FUNCTION F_InitializePolarIIChamberServiceStatus : BOOL
VAR_IN_OUT
	ServiceStatus : ST_PolarIIChamber_ServiceStatus;
END_VAR

MEMSET(ADR(ServiceStatus), 0, SIZEOF(ServiceStatus));

// Chamber
F_SetPolarIIChamberServiceIdentity(Status := ServiceStatus.Chamber.SetMode, ServiceId := E_PolarIIChamber_ServiceId.Chamber_SetMode, CompletionBehavior := E_ServiceCompletionBehavior.NaturalCompletion);
F_SetPolarIIChamberServiceIdentity(Status := ServiceStatus.Chamber.Initial, ServiceId := E_PolarIIChamber_ServiceId.Chamber_Initial, CompletionBehavior := E_ServiceCompletionBehavior.NaturalCompletion);
F_SetPolarIIChamberServiceIdentity(Status := ServiceStatus.Chamber.SingleProcess, ServiceId := E_PolarIIChamber_ServiceId.Chamber_SingleProcess, CompletionBehavior := E_ServiceCompletionBehavior.NaturalCompletion);
F_SetPolarIIChamberServiceIdentity(Status := ServiceStatus.Chamber.EMGS, ServiceId := E_PolarIIChamber_ServiceId.Chamber_EMGS, CompletionBehavior := E_ServiceCompletionBehavior.NaturalCompletion);
F_SetPolarIIChamberServiceIdentity(Status := ServiceStatus.Chamber.SetConfig, ServiceId := E_PolarIIChamber_ServiceId.Chamber_SetConfig, CompletionBehavior := E_ServiceCompletionBehavior.NaturalCompletion);
F_SetPolarIIChamberServiceIdentity(Status := ServiceStatus.Chamber.ArmAlignTest, ServiceId := E_PolarIIChamber_ServiceId.Chamber_ArmAlignTest, CompletionBehavior := E_ServiceCompletionBehavior.NaturalCompletion);
F_SetPolarIIChamberServiceIdentity(Status := ServiceStatus.Chamber.ArmTest, ServiceId := E_PolarIIChamber_ServiceId.Chamber_ArmTest, CompletionBehavior := E_ServiceCompletionBehavior.NaturalCompletion);
F_SetPolarIIChamberServiceIdentity(Status := ServiceStatus.Chamber.FlowCalibration, ServiceId := E_PolarIIChamber_ServiceId.Chamber_FlowCalibration, CompletionBehavior := E_ServiceCompletionBehavior.NaturalCompletion);
F_SetPolarIIChamberServiceIdentity(Status := ServiceStatus.Chamber.CupChamberClean, ServiceId := E_PolarIIChamber_ServiceId.Chamber_CupChamberClean, CompletionBehavior := E_ServiceCompletionBehavior.NaturalCompletion);
F_SetPolarIIChamberServiceIdentity(Status := ServiceStatus.Chamber.DoNozzleClean, ServiceId := E_PolarIIChamber_ServiceId.Chamber_DoNozzleClean, CompletionBehavior := E_ServiceCompletionBehavior.NaturalCompletion);
F_SetPolarIIChamberServiceIdentity(Status := ServiceStatus.Chamber.DoNozzlePreflush, ServiceId := E_PolarIIChamber_ServiceId.Chamber_DoNozzlePreflush, CompletionBehavior := E_ServiceCompletionBehavior.NaturalCompletion);

// Arm
F_SetPolarIIChamberServiceIdentity(Status := ServiceStatus.Arm[1].Lift.TopPos, ServiceId := E_PolarIIChamber_ServiceId.Arm1_Lift_TopPos, CompletionBehavior := E_ServiceCompletionBehavior.NaturalCompletion);
F_SetPolarIIChamberServiceIdentity(Status := ServiceStatus.Arm[1].Lift.DownPos, ServiceId := E_PolarIIChamber_ServiceId.Arm1_Lift_DownPos, CompletionBehavior := E_ServiceCompletionBehavior.NaturalCompletion);
F_SetPolarIIChamberServiceIdentity(Status := ServiceStatus.Arm[1].Rotate.JogPositive, ServiceId := E_PolarIIChamber_ServiceId.Arm1_Rotate_JogPositive, CompletionBehavior := E_ServiceCompletionBehavior.ExecuteUntilExternalStop);
F_SetPolarIIChamberServiceIdentity(Status := ServiceStatus.Arm[1].Rotate.JogNegative, ServiceId := E_PolarIIChamber_ServiceId.Arm1_Rotate_JogNegative, CompletionBehavior := E_ServiceCompletionBehavior.ExecuteUntilExternalStop);
F_SetPolarIIChamberServiceIdentity(Status := ServiceStatus.Arm[1].Rotate.IncrementalJog, ServiceId := E_PolarIIChamber_ServiceId.Arm1_Rotate_IncrementalJog, CompletionBehavior := E_ServiceCompletionBehavior.NaturalCompletion);
F_SetPolarIIChamberServiceIdentity(Status := ServiceStatus.Arm[1].Rotate.MoveRecipe, ServiceId := E_PolarIIChamber_ServiceId.Arm1_Rotate_MoveRecipe, CompletionBehavior := E_ServiceCompletionBehavior.NaturalCompletion);
F_SetPolarIIChamberServiceIdentity(Status := ServiceStatus.Arm[1].Rotate.NegLimitPos, ServiceId := E_PolarIIChamber_ServiceId.Arm1_Rotate_NegLimitPos, CompletionBehavior := E_ServiceCompletionBehavior.NaturalCompletion);
F_SetPolarIIChamberServiceIdentity(Status := ServiceStatus.Arm[1].Rotate.PosLimitPos, ServiceId := E_PolarIIChamber_ServiceId.Arm1_Rotate_PosLimitPos, CompletionBehavior := E_ServiceCompletionBehavior.NaturalCompletion);
F_SetPolarIIChamberServiceIdentity(Status := ServiceStatus.Arm[1].Rotate.NozzlePortPos, ServiceId := E_PolarIIChamber_ServiceId.Arm1_Rotate_NozPortPos, CompletionBehavior := E_ServiceCompletionBehavior.NaturalCompletion);
F_SetPolarIIChamberServiceIdentity(Status := ServiceStatus.Arm[1].Rotate.Noz1CenterPos, ServiceId := E_PolarIIChamber_ServiceId.Arm1_Rotate_Noz1CenterPos, CompletionBehavior := E_ServiceCompletionBehavior.NaturalCompletion);
F_SetPolarIIChamberServiceIdentity(Status := ServiceStatus.Arm[1].Rotate.Noz2CenterPos, ServiceId := E_PolarIIChamber_ServiceId.Arm1_Rotate_Noz2CenterPos, CompletionBehavior := E_ServiceCompletionBehavior.NaturalCompletion);
F_SetPolarIIChamberServiceIdentity(Status := ServiceStatus.Arm[1].Rotate.Noz3CenterPos, ServiceId := E_PolarIIChamber_ServiceId.Arm1_Rotate_Noz3CenterPos, CompletionBehavior := E_ServiceCompletionBehavior.NaturalCompletion);
F_SetPolarIIChamberServiceIdentity(Status := ServiceStatus.Arm[1].Nozzle[1].ChemicalSupply, ServiceId := E_PolarIIChamber_ServiceId.Arm1_Noz1_ChemicalSupply, CompletionBehavior := E_ServiceCompletionBehavior.ExecuteUntilExternalStop);
F_SetPolarIIChamberServiceIdentity(Status := ServiceStatus.Arm[1].Nozzle[2].ChemicalSupply, ServiceId := E_PolarIIChamber_ServiceId.Arm1_Noz2_ChemicalSupply, CompletionBehavior := E_ServiceCompletionBehavior.ExecuteUntilExternalStop);
F_SetPolarIIChamberServiceIdentity(Status := ServiceStatus.Arm[1].Nozzle[3].ChemicalSupply, ServiceId := E_PolarIIChamber_ServiceId.Arm1_Noz3_ChemicalSupply, CompletionBehavior := E_ServiceCompletionBehavior.ExecuteUntilExternalStop);
F_SetPolarIIChamberServiceIdentity(Status := ServiceStatus.Arm[1].NozzlePort.Nozzle[1].Supply, ServiceId := E_PolarIIChamber_ServiceId.Arm1_NozPortNoz1_Supply, CompletionBehavior := E_ServiceCompletionBehavior.ExecuteUntilExternalStop);
F_SetPolarIIChamberServiceIdentity(Status := ServiceStatus.Arm[1].NozzlePort.Nozzle[2].Supply, ServiceId := E_PolarIIChamber_ServiceId.Arm1_NozPortNoz2_Supply, CompletionBehavior := E_ServiceCompletionBehavior.ExecuteUntilExternalStop);
F_SetPolarIIChamberServiceIdentity(Status := ServiceStatus.Arm[1].NozzlePort.Nozzle[3].Supply, ServiceId := E_PolarIIChamber_ServiceId.Arm1_NozPortNoz3_Supply, CompletionBehavior := E_ServiceCompletionBehavior.ExecuteUntilExternalStop);
F_SetPolarIIChamberServiceIdentity(Status := ServiceStatus.Arm[1].NozzlePort.DrainSelect1, ServiceId := E_PolarIIChamber_ServiceId.Arm1_NozPortDrainer_Select1, CompletionBehavior := E_ServiceCompletionBehavior.NaturalCompletion);
F_SetPolarIIChamberServiceIdentity(Status := ServiceStatus.Arm[1].NozzlePort.DrainSelect2, ServiceId := E_PolarIIChamber_ServiceId.Arm1_NozPortDrainer_Select2, CompletionBehavior := E_ServiceCompletionBehavior.NaturalCompletion);
F_SetPolarIIChamberServiceIdentity(Status := ServiceStatus.Arm[1].NozzlePort.DrainSelect3, ServiceId := E_PolarIIChamber_ServiceId.Arm1_NozPortDrainer_Select3, CompletionBehavior := E_ServiceCompletionBehavior.NaturalCompletion);
F_SetPolarIIChamberServiceIdentity(Status := ServiceStatus.Arm[2].Lift.TopPos, ServiceId := E_PolarIIChamber_ServiceId.Arm2_Lift_TopPos, CompletionBehavior := E_ServiceCompletionBehavior.NaturalCompletion);
F_SetPolarIIChamberServiceIdentity(Status := ServiceStatus.Arm[2].Lift.DownPos, ServiceId := E_PolarIIChamber_ServiceId.Arm2_Lift_DownPos, CompletionBehavior := E_ServiceCompletionBehavior.NaturalCompletion);
F_SetPolarIIChamberServiceIdentity(Status := ServiceStatus.Arm[2].Rotate.JogPositive, ServiceId := E_PolarIIChamber_ServiceId.Arm2_Rotate_JogPositive, CompletionBehavior := E_ServiceCompletionBehavior.ExecuteUntilExternalStop);
F_SetPolarIIChamberServiceIdentity(Status := ServiceStatus.Arm[2].Rotate.JogNegative, ServiceId := E_PolarIIChamber_ServiceId.Arm2_Rotate_JogNegative, CompletionBehavior := E_ServiceCompletionBehavior.ExecuteUntilExternalStop);
F_SetPolarIIChamberServiceIdentity(Status := ServiceStatus.Arm[2].Rotate.IncrementalJog, ServiceId := E_PolarIIChamber_ServiceId.Arm2_Rotate_IncrementalJog, CompletionBehavior := E_ServiceCompletionBehavior.NaturalCompletion);
F_SetPolarIIChamberServiceIdentity(Status := ServiceStatus.Arm[2].Rotate.MoveRecipe, ServiceId := E_PolarIIChamber_ServiceId.Arm2_Rotate_MoveRecipe, CompletionBehavior := E_ServiceCompletionBehavior.NaturalCompletion);
F_SetPolarIIChamberServiceIdentity(Status := ServiceStatus.Arm[2].Rotate.NegLimitPos, ServiceId := E_PolarIIChamber_ServiceId.Arm2_Rotate_NegLimitPos, CompletionBehavior := E_ServiceCompletionBehavior.NaturalCompletion);
F_SetPolarIIChamberServiceIdentity(Status := ServiceStatus.Arm[2].Rotate.PosLimitPos, ServiceId := E_PolarIIChamber_ServiceId.Arm2_Rotate_PosLimitPos, CompletionBehavior := E_ServiceCompletionBehavior.NaturalCompletion);
F_SetPolarIIChamberServiceIdentity(Status := ServiceStatus.Arm[2].Rotate.NozzlePortPos, ServiceId := E_PolarIIChamber_ServiceId.Arm2_Rotate_NozPortPos, CompletionBehavior := E_ServiceCompletionBehavior.NaturalCompletion);
F_SetPolarIIChamberServiceIdentity(Status := ServiceStatus.Arm[2].Rotate.Noz1CenterPos, ServiceId := E_PolarIIChamber_ServiceId.Arm2_Rotate_Noz1CenterPos, CompletionBehavior := E_ServiceCompletionBehavior.NaturalCompletion);
F_SetPolarIIChamberServiceIdentity(Status := ServiceStatus.Arm[2].Rotate.Noz2CenterPos, ServiceId := E_PolarIIChamber_ServiceId.Arm2_Rotate_Noz2CenterPos, CompletionBehavior := E_ServiceCompletionBehavior.NaturalCompletion);
F_SetPolarIIChamberServiceIdentity(Status := ServiceStatus.Arm[2].Rotate.Noz3CenterPos, ServiceId := E_PolarIIChamber_ServiceId.Arm2_Rotate_Noz3CenterPos, CompletionBehavior := E_ServiceCompletionBehavior.NaturalCompletion);
F_SetPolarIIChamberServiceIdentity(Status := ServiceStatus.Arm[2].Nozzle[1].ChemicalSupply, ServiceId := E_PolarIIChamber_ServiceId.Arm2_Noz1_ChemicalSupply, CompletionBehavior := E_ServiceCompletionBehavior.ExecuteUntilExternalStop);
F_SetPolarIIChamberServiceIdentity(Status := ServiceStatus.Arm[2].Nozzle[2].ChemicalSupply, ServiceId := E_PolarIIChamber_ServiceId.Arm2_Noz2_ChemicalSupply, CompletionBehavior := E_ServiceCompletionBehavior.ExecuteUntilExternalStop);
F_SetPolarIIChamberServiceIdentity(Status := ServiceStatus.Arm[2].Nozzle[3].ChemicalSupply, ServiceId := E_PolarIIChamber_ServiceId.Arm2_Noz3_ChemicalSupply, CompletionBehavior := E_ServiceCompletionBehavior.ExecuteUntilExternalStop);
F_SetPolarIIChamberServiceIdentity(Status := ServiceStatus.Arm[2].NozzlePort.Nozzle[1].Supply, ServiceId := E_PolarIIChamber_ServiceId.Arm2_NozPortNoz1_Supply, CompletionBehavior := E_ServiceCompletionBehavior.ExecuteUntilExternalStop);
F_SetPolarIIChamberServiceIdentity(Status := ServiceStatus.Arm[2].NozzlePort.Nozzle[2].Supply, ServiceId := E_PolarIIChamber_ServiceId.Arm2_NozPortNoz2_Supply, CompletionBehavior := E_ServiceCompletionBehavior.ExecuteUntilExternalStop);
F_SetPolarIIChamberServiceIdentity(Status := ServiceStatus.Arm[2].NozzlePort.Nozzle[3].Supply, ServiceId := E_PolarIIChamber_ServiceId.Arm2_NozPortNoz3_Supply, CompletionBehavior := E_ServiceCompletionBehavior.ExecuteUntilExternalStop);
F_SetPolarIIChamberServiceIdentity(Status := ServiceStatus.Arm[2].NozzlePort.DrainSelect1, ServiceId := E_PolarIIChamber_ServiceId.Arm2_NozPortDrainer_Select1, CompletionBehavior := E_ServiceCompletionBehavior.NaturalCompletion);
F_SetPolarIIChamberServiceIdentity(Status := ServiceStatus.Arm[2].NozzlePort.DrainSelect2, ServiceId := E_PolarIIChamber_ServiceId.Arm2_NozPortDrainer_Select2, CompletionBehavior := E_ServiceCompletionBehavior.NaturalCompletion);
F_SetPolarIIChamberServiceIdentity(Status := ServiceStatus.Arm[2].NozzlePort.DrainSelect3, ServiceId := E_PolarIIChamber_ServiceId.Arm2_NozPortDrainer_Select3, CompletionBehavior := E_ServiceCompletionBehavior.NaturalCompletion);
F_SetPolarIIChamberServiceIdentity(Status := ServiceStatus.Arm[3].Lift.TopPos, ServiceId := E_PolarIIChamber_ServiceId.Arm3_Lift_TopPos, CompletionBehavior := E_ServiceCompletionBehavior.NaturalCompletion);
F_SetPolarIIChamberServiceIdentity(Status := ServiceStatus.Arm[3].Lift.DownPos, ServiceId := E_PolarIIChamber_ServiceId.Arm3_Lift_DownPos, CompletionBehavior := E_ServiceCompletionBehavior.NaturalCompletion);
F_SetPolarIIChamberServiceIdentity(Status := ServiceStatus.Arm[3].Rotate.JogPositive, ServiceId := E_PolarIIChamber_ServiceId.Arm3_Rotate_JogPositive, CompletionBehavior := E_ServiceCompletionBehavior.ExecuteUntilExternalStop);
F_SetPolarIIChamberServiceIdentity(Status := ServiceStatus.Arm[3].Rotate.JogNegative, ServiceId := E_PolarIIChamber_ServiceId.Arm3_Rotate_JogNegative, CompletionBehavior := E_ServiceCompletionBehavior.ExecuteUntilExternalStop);
F_SetPolarIIChamberServiceIdentity(Status := ServiceStatus.Arm[3].Rotate.IncrementalJog, ServiceId := E_PolarIIChamber_ServiceId.Arm3_Rotate_IncrementalJog, CompletionBehavior := E_ServiceCompletionBehavior.NaturalCompletion);
F_SetPolarIIChamberServiceIdentity(Status := ServiceStatus.Arm[3].Rotate.MoveRecipe, ServiceId := E_PolarIIChamber_ServiceId.Arm3_Rotate_MoveRecipe, CompletionBehavior := E_ServiceCompletionBehavior.NaturalCompletion);
F_SetPolarIIChamberServiceIdentity(Status := ServiceStatus.Arm[3].Rotate.NegLimitPos, ServiceId := E_PolarIIChamber_ServiceId.Arm3_Rotate_NegLimitPos, CompletionBehavior := E_ServiceCompletionBehavior.NaturalCompletion);
F_SetPolarIIChamberServiceIdentity(Status := ServiceStatus.Arm[3].Rotate.PosLimitPos, ServiceId := E_PolarIIChamber_ServiceId.Arm3_Rotate_PosLimitPos, CompletionBehavior := E_ServiceCompletionBehavior.NaturalCompletion);
F_SetPolarIIChamberServiceIdentity(Status := ServiceStatus.Arm[3].Rotate.Noz1CenterPos, ServiceId := E_PolarIIChamber_ServiceId.Arm3_Rotate_Noz1CenterPos, CompletionBehavior := E_ServiceCompletionBehavior.NaturalCompletion);
F_SetPolarIIChamberServiceIdentity(Status := ServiceStatus.Arm[3].Rotate.Noz2CenterPos, ServiceId := E_PolarIIChamber_ServiceId.Arm3_Rotate_Noz2CenterPos, CompletionBehavior := E_ServiceCompletionBehavior.NaturalCompletion);
F_SetPolarIIChamberServiceIdentity(Status := ServiceStatus.Arm[3].Nozzle[1].ChemicalSupply, ServiceId := E_PolarIIChamber_ServiceId.Arm3_Noz1_ChemicalSupply, CompletionBehavior := E_ServiceCompletionBehavior.ExecuteUntilExternalStop);
F_SetPolarIIChamberServiceIdentity(Status := ServiceStatus.Arm[3].Nozzle[2].ChemicalSupply, ServiceId := E_PolarIIChamber_ServiceId.Arm3_Noz2_ChemicalSupply, CompletionBehavior := E_ServiceCompletionBehavior.ExecuteUntilExternalStop);
// Arm[3] has no third nozzle or nozzle port. Keep ServiceId = 0, but provide
// CompletionBehavior so the current SDK STRUCT scanner can complete validation.
ServiceStatus.Arm[3].Rotate.NozzlePortPos.CompletionBehavior := E_ServiceCompletionBehavior.NaturalCompletion;
ServiceStatus.Arm[3].Rotate.Noz3CenterPos.CompletionBehavior := E_ServiceCompletionBehavior.NaturalCompletion;
ServiceStatus.Arm[3].Nozzle[3].ChemicalSupply.CompletionBehavior := E_ServiceCompletionBehavior.ExecuteUntilExternalStop;
ServiceStatus.Arm[3].NozzlePort.Nozzle[1].Supply.CompletionBehavior := E_ServiceCompletionBehavior.ExecuteUntilExternalStop;
ServiceStatus.Arm[3].NozzlePort.Nozzle[2].Supply.CompletionBehavior := E_ServiceCompletionBehavior.ExecuteUntilExternalStop;
ServiceStatus.Arm[3].NozzlePort.Nozzle[3].Supply.CompletionBehavior := E_ServiceCompletionBehavior.ExecuteUntilExternalStop;
ServiceStatus.Arm[3].NozzlePort.DrainSelect1.CompletionBehavior := E_ServiceCompletionBehavior.NaturalCompletion;
ServiceStatus.Arm[3].NozzlePort.DrainSelect2.CompletionBehavior := E_ServiceCompletionBehavior.NaturalCompletion;
ServiceStatus.Arm[3].NozzlePort.DrainSelect3.CompletionBehavior := E_ServiceCompletionBehavior.NaturalCompletion;
F_SetPolarIIChamberServiceIdentity(Status := ServiceStatus.Arm[4].Lift.TopPos, ServiceId := E_PolarIIChamber_ServiceId.Arm4_Lift_TopPos, CompletionBehavior := E_ServiceCompletionBehavior.NaturalCompletion);
F_SetPolarIIChamberServiceIdentity(Status := ServiceStatus.Arm[4].Lift.DownPos, ServiceId := E_PolarIIChamber_ServiceId.Arm4_Lift_DownPos, CompletionBehavior := E_ServiceCompletionBehavior.NaturalCompletion);
F_SetPolarIIChamberServiceIdentity(Status := ServiceStatus.Arm[4].Rotate.JogPositive, ServiceId := E_PolarIIChamber_ServiceId.Arm4_Rotate_JogPositive, CompletionBehavior := E_ServiceCompletionBehavior.ExecuteUntilExternalStop);
F_SetPolarIIChamberServiceIdentity(Status := ServiceStatus.Arm[4].Rotate.JogNegative, ServiceId := E_PolarIIChamber_ServiceId.Arm4_Rotate_JogNegative, CompletionBehavior := E_ServiceCompletionBehavior.ExecuteUntilExternalStop);
F_SetPolarIIChamberServiceIdentity(Status := ServiceStatus.Arm[4].Rotate.IncrementalJog, ServiceId := E_PolarIIChamber_ServiceId.Arm4_Rotate_IncrementalJog, CompletionBehavior := E_ServiceCompletionBehavior.NaturalCompletion);
F_SetPolarIIChamberServiceIdentity(Status := ServiceStatus.Arm[4].Rotate.MoveRecipe, ServiceId := E_PolarIIChamber_ServiceId.Arm4_Rotate_MoveRecipe, CompletionBehavior := E_ServiceCompletionBehavior.NaturalCompletion);
F_SetPolarIIChamberServiceIdentity(Status := ServiceStatus.Arm[4].Rotate.NegLimitPos, ServiceId := E_PolarIIChamber_ServiceId.Arm4_Rotate_NegLimitPos, CompletionBehavior := E_ServiceCompletionBehavior.NaturalCompletion);
F_SetPolarIIChamberServiceIdentity(Status := ServiceStatus.Arm[4].Rotate.PosLimitPos, ServiceId := E_PolarIIChamber_ServiceId.Arm4_Rotate_PosLimitPos, CompletionBehavior := E_ServiceCompletionBehavior.NaturalCompletion);
F_SetPolarIIChamberServiceIdentity(Status := ServiceStatus.Arm[4].Rotate.Noz1CenterPos, ServiceId := E_PolarIIChamber_ServiceId.Arm4_Rotate_Noz1CenterPos, CompletionBehavior := E_ServiceCompletionBehavior.NaturalCompletion);
F_SetPolarIIChamberServiceIdentity(Status := ServiceStatus.Arm[4].Nozzle[1].ChemicalSupply, ServiceId := E_PolarIIChamber_ServiceId.Arm4_Noz1_ChemicalSupply, CompletionBehavior := E_ServiceCompletionBehavior.ExecuteUntilExternalStop);
// Arm[4] has no second/third nozzle or nozzle port. Keep ServiceId = 0, but
// provide CompletionBehavior for compatibility with the current SDK scanner.
ServiceStatus.Arm[4].Rotate.NozzlePortPos.CompletionBehavior := E_ServiceCompletionBehavior.NaturalCompletion;
ServiceStatus.Arm[4].Rotate.Noz2CenterPos.CompletionBehavior := E_ServiceCompletionBehavior.NaturalCompletion;
ServiceStatus.Arm[4].Rotate.Noz3CenterPos.CompletionBehavior := E_ServiceCompletionBehavior.NaturalCompletion;
ServiceStatus.Arm[4].Nozzle[2].ChemicalSupply.CompletionBehavior := E_ServiceCompletionBehavior.ExecuteUntilExternalStop;
ServiceStatus.Arm[4].Nozzle[3].ChemicalSupply.CompletionBehavior := E_ServiceCompletionBehavior.ExecuteUntilExternalStop;
ServiceStatus.Arm[4].NozzlePort.Nozzle[1].Supply.CompletionBehavior := E_ServiceCompletionBehavior.ExecuteUntilExternalStop;
ServiceStatus.Arm[4].NozzlePort.Nozzle[2].Supply.CompletionBehavior := E_ServiceCompletionBehavior.ExecuteUntilExternalStop;
ServiceStatus.Arm[4].NozzlePort.Nozzle[3].Supply.CompletionBehavior := E_ServiceCompletionBehavior.ExecuteUntilExternalStop;
ServiceStatus.Arm[4].NozzlePort.DrainSelect1.CompletionBehavior := E_ServiceCompletionBehavior.NaturalCompletion;
ServiceStatus.Arm[4].NozzlePort.DrainSelect2.CompletionBehavior := E_ServiceCompletionBehavior.NaturalCompletion;
ServiceStatus.Arm[4].NozzlePort.DrainSelect3.CompletionBehavior := E_ServiceCompletionBehavior.NaturalCompletion;

// Cup
F_SetPolarIIChamberServiceIdentity(Status := ServiceStatus.Cup[1].Lift.JogPositive, ServiceId := E_PolarIIChamber_ServiceId.Cup1_Lift_JogPositive, CompletionBehavior := E_ServiceCompletionBehavior.ExecuteUntilExternalStop);
F_SetPolarIIChamberServiceIdentity(Status := ServiceStatus.Cup[1].Lift.JogNegative, ServiceId := E_PolarIIChamber_ServiceId.Cup1_Lift_JogNegative, CompletionBehavior := E_ServiceCompletionBehavior.ExecuteUntilExternalStop);
F_SetPolarIIChamberServiceIdentity(Status := ServiceStatus.Cup[1].Lift.IncrementalJog, ServiceId := E_PolarIIChamber_ServiceId.Cup1_Lift_IncrementalJog, CompletionBehavior := E_ServiceCompletionBehavior.NaturalCompletion);
F_SetPolarIIChamberServiceIdentity(Status := ServiceStatus.Cup[1].Lift.DecoupleStop, ServiceId := E_PolarIIChamber_ServiceId.Cup1_Lift_DecoupleStop, CompletionBehavior := E_ServiceCompletionBehavior.NaturalCompletion);
F_SetPolarIIChamberServiceIdentity(Status := ServiceStatus.Cup[1].Lift.TopPos, ServiceId := E_PolarIIChamber_ServiceId.Cup1_Lift_TopPos, CompletionBehavior := E_ServiceCompletionBehavior.NaturalCompletion);
F_SetPolarIIChamberServiceIdentity(Status := ServiceStatus.Cup[1].Lift.MiddlePos, ServiceId := E_PolarIIChamber_ServiceId.Cup1_Lift_MiddlePos, CompletionBehavior := E_ServiceCompletionBehavior.NaturalCompletion);
F_SetPolarIIChamberServiceIdentity(Status := ServiceStatus.Cup[1].Lift.DownPos, ServiceId := E_PolarIIChamber_ServiceId.Cup1_Lift_DownPos, CompletionBehavior := E_ServiceCompletionBehavior.NaturalCompletion);
F_SetPolarIIChamberServiceIdentity(Status := ServiceStatus.Cup[1].Drainer.Select1, ServiceId := E_PolarIIChamber_ServiceId.Cup1_Drainer_Select1, CompletionBehavior := E_ServiceCompletionBehavior.NaturalCompletion);
F_SetPolarIIChamberServiceIdentity(Status := ServiceStatus.Cup[1].Drainer.Select2, ServiceId := E_PolarIIChamber_ServiceId.Cup1_Drainer_Select2, CompletionBehavior := E_ServiceCompletionBehavior.NaturalCompletion);
F_SetPolarIIChamberServiceIdentity(Status := ServiceStatus.Cup[1].Drainer.Select3, ServiceId := E_PolarIIChamber_ServiceId.Cup1_Drainer_Select3, CompletionBehavior := E_ServiceCompletionBehavior.NaturalCompletion);
F_SetPolarIIChamberServiceIdentity(Status := ServiceStatus.Cup[2].Lift.JogPositive, ServiceId := E_PolarIIChamber_ServiceId.Cup2_Lift_JogPositive, CompletionBehavior := E_ServiceCompletionBehavior.ExecuteUntilExternalStop);
F_SetPolarIIChamberServiceIdentity(Status := ServiceStatus.Cup[2].Lift.JogNegative, ServiceId := E_PolarIIChamber_ServiceId.Cup2_Lift_JogNegative, CompletionBehavior := E_ServiceCompletionBehavior.ExecuteUntilExternalStop);
F_SetPolarIIChamberServiceIdentity(Status := ServiceStatus.Cup[2].Lift.IncrementalJog, ServiceId := E_PolarIIChamber_ServiceId.Cup2_Lift_IncrementalJog, CompletionBehavior := E_ServiceCompletionBehavior.NaturalCompletion);
F_SetPolarIIChamberServiceIdentity(Status := ServiceStatus.Cup[2].Lift.DecoupleStop, ServiceId := E_PolarIIChamber_ServiceId.Cup2_Lift_DecoupleStop, CompletionBehavior := E_ServiceCompletionBehavior.NaturalCompletion);
F_SetPolarIIChamberServiceIdentity(Status := ServiceStatus.Cup[2].Lift.TopPos, ServiceId := E_PolarIIChamber_ServiceId.Cup2_Lift_TopPos, CompletionBehavior := E_ServiceCompletionBehavior.NaturalCompletion);
F_SetPolarIIChamberServiceIdentity(Status := ServiceStatus.Cup[2].Lift.MiddlePos, ServiceId := E_PolarIIChamber_ServiceId.Cup2_Lift_MiddlePos, CompletionBehavior := E_ServiceCompletionBehavior.NaturalCompletion);
F_SetPolarIIChamberServiceIdentity(Status := ServiceStatus.Cup[2].Lift.DownPos, ServiceId := E_PolarIIChamber_ServiceId.Cup2_Lift_DownPos, CompletionBehavior := E_ServiceCompletionBehavior.NaturalCompletion);
F_SetPolarIIChamberServiceIdentity(Status := ServiceStatus.Cup[2].Drainer.Select1, ServiceId := E_PolarIIChamber_ServiceId.Cup2_Drainer_Select1, CompletionBehavior := E_ServiceCompletionBehavior.NaturalCompletion);
F_SetPolarIIChamberServiceIdentity(Status := ServiceStatus.Cup[2].Drainer.Select2, ServiceId := E_PolarIIChamber_ServiceId.Cup2_Drainer_Select2, CompletionBehavior := E_ServiceCompletionBehavior.NaturalCompletion);
F_SetPolarIIChamberServiceIdentity(Status := ServiceStatus.Cup[2].Drainer.Select3, ServiceId := E_PolarIIChamber_ServiceId.Cup2_Drainer_Select3, CompletionBehavior := E_ServiceCompletionBehavior.NaturalCompletion);
F_SetPolarIIChamberServiceIdentity(Status := ServiceStatus.Cup[3].Lift.JogPositive, ServiceId := E_PolarIIChamber_ServiceId.Cup3_Lift_JogPositive, CompletionBehavior := E_ServiceCompletionBehavior.ExecuteUntilExternalStop);
F_SetPolarIIChamberServiceIdentity(Status := ServiceStatus.Cup[3].Lift.JogNegative, ServiceId := E_PolarIIChamber_ServiceId.Cup3_Lift_JogNegative, CompletionBehavior := E_ServiceCompletionBehavior.ExecuteUntilExternalStop);
F_SetPolarIIChamberServiceIdentity(Status := ServiceStatus.Cup[3].Lift.IncrementalJog, ServiceId := E_PolarIIChamber_ServiceId.Cup3_Lift_IncrementalJog, CompletionBehavior := E_ServiceCompletionBehavior.NaturalCompletion);
F_SetPolarIIChamberServiceIdentity(Status := ServiceStatus.Cup[3].Lift.DecoupleStop, ServiceId := E_PolarIIChamber_ServiceId.Cup3_Lift_DecoupleStop, CompletionBehavior := E_ServiceCompletionBehavior.NaturalCompletion);
F_SetPolarIIChamberServiceIdentity(Status := ServiceStatus.Cup[3].Lift.TopPos, ServiceId := E_PolarIIChamber_ServiceId.Cup3_Lift_TopPos, CompletionBehavior := E_ServiceCompletionBehavior.NaturalCompletion);
F_SetPolarIIChamberServiceIdentity(Status := ServiceStatus.Cup[3].Lift.MiddlePos, ServiceId := E_PolarIIChamber_ServiceId.Cup3_Lift_MiddlePos, CompletionBehavior := E_ServiceCompletionBehavior.NaturalCompletion);
F_SetPolarIIChamberServiceIdentity(Status := ServiceStatus.Cup[3].Lift.DownPos, ServiceId := E_PolarIIChamber_ServiceId.Cup3_Lift_DownPos, CompletionBehavior := E_ServiceCompletionBehavior.NaturalCompletion);
F_SetPolarIIChamberServiceIdentity(Status := ServiceStatus.Cup[3].Drainer.Select1, ServiceId := E_PolarIIChamber_ServiceId.Cup3_Drainer_Select1, CompletionBehavior := E_ServiceCompletionBehavior.NaturalCompletion);
F_SetPolarIIChamberServiceIdentity(Status := ServiceStatus.Cup[3].Drainer.Select2, ServiceId := E_PolarIIChamber_ServiceId.Cup3_Drainer_Select2, CompletionBehavior := E_ServiceCompletionBehavior.NaturalCompletion);
F_SetPolarIIChamberServiceIdentity(Status := ServiceStatus.Cup[3].Drainer.Select3, ServiceId := E_PolarIIChamber_ServiceId.Cup3_Drainer_Select3, CompletionBehavior := E_ServiceCompletionBehavior.NaturalCompletion);
F_SetPolarIIChamberServiceIdentity(Status := ServiceStatus.Cup[4].Lift.JogPositive, ServiceId := E_PolarIIChamber_ServiceId.Cup4_Lift_JogPositive, CompletionBehavior := E_ServiceCompletionBehavior.ExecuteUntilExternalStop);
F_SetPolarIIChamberServiceIdentity(Status := ServiceStatus.Cup[4].Lift.JogNegative, ServiceId := E_PolarIIChamber_ServiceId.Cup4_Lift_JogNegative, CompletionBehavior := E_ServiceCompletionBehavior.ExecuteUntilExternalStop);
F_SetPolarIIChamberServiceIdentity(Status := ServiceStatus.Cup[4].Lift.IncrementalJog, ServiceId := E_PolarIIChamber_ServiceId.Cup4_Lift_IncrementalJog, CompletionBehavior := E_ServiceCompletionBehavior.NaturalCompletion);
F_SetPolarIIChamberServiceIdentity(Status := ServiceStatus.Cup[4].Lift.DecoupleStop, ServiceId := E_PolarIIChamber_ServiceId.Cup4_Lift_DecoupleStop, CompletionBehavior := E_ServiceCompletionBehavior.NaturalCompletion);
F_SetPolarIIChamberServiceIdentity(Status := ServiceStatus.Cup[4].Lift.TopPos, ServiceId := E_PolarIIChamber_ServiceId.Cup4_Lift_TopPos, CompletionBehavior := E_ServiceCompletionBehavior.NaturalCompletion);
F_SetPolarIIChamberServiceIdentity(Status := ServiceStatus.Cup[4].Lift.MiddlePos, ServiceId := E_PolarIIChamber_ServiceId.Cup4_Lift_MiddlePos, CompletionBehavior := E_ServiceCompletionBehavior.NaturalCompletion);
F_SetPolarIIChamberServiceIdentity(Status := ServiceStatus.Cup[4].Lift.DownPos, ServiceId := E_PolarIIChamber_ServiceId.Cup4_Lift_DownPos, CompletionBehavior := E_ServiceCompletionBehavior.NaturalCompletion);
F_SetPolarIIChamberServiceIdentity(Status := ServiceStatus.Cup[4].Drainer.Select1, ServiceId := E_PolarIIChamber_ServiceId.Cup4_Drainer_Select1, CompletionBehavior := E_ServiceCompletionBehavior.NaturalCompletion);
F_SetPolarIIChamberServiceIdentity(Status := ServiceStatus.Cup[4].Drainer.Select2, ServiceId := E_PolarIIChamber_ServiceId.Cup4_Drainer_Select2, CompletionBehavior := E_ServiceCompletionBehavior.NaturalCompletion);
F_SetPolarIIChamberServiceIdentity(Status := ServiceStatus.Cup[4].Drainer.Select3, ServiceId := E_PolarIIChamber_ServiceId.Cup4_Drainer_Select3, CompletionBehavior := E_ServiceCompletionBehavior.NaturalCompletion);

// Holder
F_SetPolarIIChamberServiceIdentity(Status := ServiceStatus.Holder.Gripper.Open, ServiceId := E_PolarIIChamber_ServiceId.Holder_Gripper_Open, CompletionBehavior := E_ServiceCompletionBehavior.NaturalCompletion);
F_SetPolarIIChamberServiceIdentity(Status := ServiceStatus.Holder.Gripper.Close, ServiceId := E_PolarIIChamber_ServiceId.Holder_Gripper_Close, CompletionBehavior := E_ServiceCompletionBehavior.NaturalCompletion);
F_SetPolarIIChamberServiceIdentity(Status := ServiceStatus.Holder.Rotate.OPR, ServiceId := E_PolarIIChamber_ServiceId.Holder_Rotate_OPR, CompletionBehavior := E_ServiceCompletionBehavior.NaturalCompletion);
F_SetPolarIIChamberServiceIdentity(Status := ServiceStatus.Holder.Rotate.MoveVelocityCW, ServiceId := E_PolarIIChamber_ServiceId.Holder_Rotate_MoveVelocityCW, CompletionBehavior := E_ServiceCompletionBehavior.ExecuteUntilExternalStop);
F_SetPolarIIChamberServiceIdentity(Status := ServiceStatus.Holder.Rotate.MoveVelocityCCW, ServiceId := E_PolarIIChamber_ServiceId.Holder_Rotate_MoveVelocityCCW, CompletionBehavior := E_ServiceCompletionBehavior.ExecuteUntilExternalStop);
F_SetPolarIIChamberServiceIdentity(Status := ServiceStatus.Holder.Rotate.MoveModulo, ServiceId := E_PolarIIChamber_ServiceId.Holder_Rotate_MoveModulo, CompletionBehavior := E_ServiceCompletionBehavior.NaturalCompletion);
F_SetPolarIIChamberServiceIdentity(Status := ServiceStatus.Holder.VacuumEstablish, ServiceId := E_PolarIIChamber_ServiceId.Holder_VacuumEstablish, CompletionBehavior := E_ServiceCompletionBehavior.ExecuteUntilExternalStop);

// FixedNozzle
F_SetPolarIIChamberServiceIdentity(Status := ServiceStatus.FixedNozzle[1].ChemicalSupply, ServiceId := E_PolarIIChamber_ServiceId.FixedNoz1_ChemicalSupply, CompletionBehavior := E_ServiceCompletionBehavior.ExecuteUntilExternalStop);
F_SetPolarIIChamberServiceIdentity(Status := ServiceStatus.FixedNozzle[2].ChemicalSupply, ServiceId := E_PolarIIChamber_ServiceId.FixedNoz2_ChemicalSupply, CompletionBehavior := E_ServiceCompletionBehavior.ExecuteUntilExternalStop);
F_SetPolarIIChamberServiceIdentity(Status := ServiceStatus.FixedNozzle[3].ChemicalSupply, ServiceId := E_PolarIIChamber_ServiceId.FixedNoz3_ChemicalSupply, CompletionBehavior := E_ServiceCompletionBehavior.ExecuteUntilExternalStop);
F_SetPolarIIChamberServiceIdentity(Status := ServiceStatus.FixedNozzle[4].ChemicalSupply, ServiceId := E_PolarIIChamber_ServiceId.FixedNoz4_ChemicalSupply, CompletionBehavior := E_ServiceCompletionBehavior.ExecuteUntilExternalStop);

// OutsideRing
F_SetPolarIIChamberServiceIdentity(Status := ServiceStatus.OutsideRing.Lift.TopPos, ServiceId := E_PolarIIChamber_ServiceId.OutsideRing_Lift_TopPos, CompletionBehavior := E_ServiceCompletionBehavior.NaturalCompletion);
F_SetPolarIIChamberServiceIdentity(Status := ServiceStatus.OutsideRing.Lift.DownPos, ServiceId := E_PolarIIChamber_ServiceId.OutsideRing_Lift_DownPos, CompletionBehavior := E_ServiceCompletionBehavior.NaturalCompletion);
F_SetPolarIIChamberServiceIdentity(Status := ServiceStatus.OutsideRing.Rotate.MoveVelocityCW, ServiceId := E_PolarIIChamber_ServiceId.OutsideRing_Rotate_MoveVelocityCW, CompletionBehavior := E_ServiceCompletionBehavior.ExecuteUntilExternalStop);
F_SetPolarIIChamberServiceIdentity(Status := ServiceStatus.OutsideRing.Rotate.MoveVelocityCCW, ServiceId := E_PolarIIChamber_ServiceId.OutsideRing_Rotate_MoveVelocityCCW, CompletionBehavior := E_ServiceCompletionBehavior.ExecuteUntilExternalStop);

// Shutter
F_SetPolarIIChamberServiceIdentity(Status := ServiceStatus.Shutter.Open, ServiceId := E_PolarIIChamber_ServiceId.Shutter_Open, CompletionBehavior := E_ServiceCompletionBehavior.NaturalCompletion);
F_SetPolarIIChamberServiceIdentity(Status := ServiceStatus.Shutter.Close, ServiceId := E_PolarIIChamber_ServiceId.Shutter_Close, CompletionBehavior := E_ServiceCompletionBehavior.NaturalCompletion);

// Exhaust
F_SetPolarIIChamberServiceIdentity(Status := ServiceStatus.Exhaust.Fan[1].SupplyFlowPID, ServiceId := E_PolarIIChamber_ServiceId.ExhaustFan1_SupplyFlowPID, CompletionBehavior := E_ServiceCompletionBehavior.ExecuteUntilExternalStop);
F_SetPolarIIChamberServiceIdentity(Status := ServiceStatus.Exhaust.Fan[2].SupplyFlowPID, ServiceId := E_PolarIIChamber_ServiceId.ExhaustFan2_SupplyFlowPID, CompletionBehavior := E_ServiceCompletionBehavior.ExecuteUntilExternalStop);
F_SetPolarIIChamberServiceIdentity(Status := ServiceStatus.Exhaust.Fan[3].SupplyFlowPID, ServiceId := E_PolarIIChamber_ServiceId.ExhaustFan3_SupplyFlowPID, CompletionBehavior := E_ServiceCompletionBehavior.ExecuteUntilExternalStop);
F_SetPolarIIChamberServiceIdentity(Status := ServiceStatus.Exhaust.Fan[4].SupplyFlowPID, ServiceId := E_PolarIIChamber_ServiceId.ExhaustFan4_SupplyFlowPID, CompletionBehavior := E_ServiceCompletionBehavior.ExecuteUntilExternalStop);
F_SetPolarIIChamberServiceIdentity(Status := ServiceStatus.Exhaust.Damper.AEX, ServiceId := E_PolarIIChamber_ServiceId.ExhaustDamper_AEX, CompletionBehavior := E_ServiceCompletionBehavior.NaturalCompletion);
F_SetPolarIIChamberServiceIdentity(Status := ServiceStatus.Exhaust.Damper.SEX, ServiceId := E_PolarIIChamber_ServiceId.ExhaustDamper_SEX, CompletionBehavior := E_ServiceCompletionBehavior.NaturalCompletion);

// SideVent
F_SetPolarIIChamberServiceIdentity(Status := ServiceStatus.SideVent[1].Open, ServiceId := E_PolarIIChamber_ServiceId.SideVent1_Open, CompletionBehavior := E_ServiceCompletionBehavior.NaturalCompletion);
F_SetPolarIIChamberServiceIdentity(Status := ServiceStatus.SideVent[1].Close, ServiceId := E_PolarIIChamber_ServiceId.SideVent1_Close, CompletionBehavior := E_ServiceCompletionBehavior.NaturalCompletion);
F_SetPolarIIChamberServiceIdentity(Status := ServiceStatus.SideVent[2].Open, ServiceId := E_PolarIIChamber_ServiceId.SideVent2_Open, CompletionBehavior := E_ServiceCompletionBehavior.NaturalCompletion);
F_SetPolarIIChamberServiceIdentity(Status := ServiceStatus.SideVent[2].Close, ServiceId := E_PolarIIChamber_ServiceId.SideVent2_Close, CompletionBehavior := E_ServiceCompletionBehavior.NaturalCompletion);
F_SetPolarIIChamberServiceIdentity(Status := ServiceStatus.SideVent[3].Open, ServiceId := E_PolarIIChamber_ServiceId.SideVent3_Open, CompletionBehavior := E_ServiceCompletionBehavior.NaturalCompletion);
F_SetPolarIIChamberServiceIdentity(Status := ServiceStatus.SideVent[3].Close, ServiceId := E_PolarIIChamber_ServiceId.SideVent3_Close, CompletionBehavior := E_ServiceCompletionBehavior.NaturalCompletion);
F_SetPolarIIChamberServiceIdentity(Status := ServiceStatus.SideVent[4].Open, ServiceId := E_PolarIIChamber_ServiceId.SideVent4_Open, CompletionBehavior := E_ServiceCompletionBehavior.NaturalCompletion);
F_SetPolarIIChamberServiceIdentity(Status := ServiceStatus.SideVent[4].Close, ServiceId := E_PolarIIChamber_ServiceId.SideVent4_Close, CompletionBehavior := E_ServiceCompletionBehavior.NaturalCompletion);

F_InitializePolarIIChamberServiceStatus := TRUE;

END_FUNCTION

(* stored: Version 1.1.0.1, ProductVersion 3.1.4026.26
   POU F_InitializePolarIIChamberServiceStatus: Id {a9ad0d91-5e87-4198-bb35-bce6689b1002}, SpecialFunc None *)
